(* IEC 61131-3 sources: Jacob-Formschaumtechnik-ISEL-CNC-Retrofit/twincat/PLC/src/1_IO, 3 files *)

(* ---- ST_AxisDrive.st ---- *)
(* Generische Achsschnittstelle. Die Maschinenlogik kennt nur diese Struktur.
   Die Zuordnung zu Klemmen/PDOs erfolgt ausschliesslich in FB_AxisMap_*. *)
TYPE ST_AxisDrive :
STRUCT
    (* Kommando (Logik -> Antrieb) *)
    bEnableReq   : BOOL;   (* Reglerfreigabe angefordert; wirkt nur mit Sicherheitsfreigabe *)
    bResetReq    : BOOL;
    (* Status (Antrieb -> Logik) *)
    bReady       : BOOL;
    bEnabled     : BOOL;
    bFault       : BOOL;
    nFaultCode   : UDINT;
    bHomed       : BOOL;
    bHwLimitPlus : BOOL;   (* Endschalter, Ruhestrom: FALSE = ausgeloest *)
    bHwLimitMinus: BOOL;
    rActPos      : LREAL;  (* mm *)
    rFollowErr   : LREAL;  (* mm *)
END_STRUCT
END_TYPE

(* ---- FB_AxisMap_Canopen.st ---- *)
(* Variante A: CANopen DS402 ueber EL6751. NOCH NICHT IMPLEMENTIERT.
   Wartet auf: Bestaetigung iMD 40 im Interpolated Position Mode mit TwinCAT CNC,
   PDO-Zuordnung und Achsnummern (Schaltplan fehlt). Die Logik darf diesen Baustein
   nicht direkt kennen, nur ST_AxisDrive. *)
FUNCTION_BLOCK FB_AxisMap_Canopen
VAR_INPUT
    bSafeEnable : BOOL;
END_VAR
VAR_IN_OUT
    stAxis : ST_AxisDrive;
END_VAR

(* [offen] Zuordnung der Prozessdaten *)
stAxis.bReady   := FALSE;
stAxis.bEnabled := FALSE;
stAxis.bFault   := TRUE;
stAxis.nFaultCode := 16#FFFF0001;  (* nicht implementiert: Maschine bleibt gesperrt *)
END_FUNCTION_BLOCK

(* ---- FB_AxisMap_Simulation.st ---- *)
(* Simulationsabbild fuer Usermode Runtime ohne Hardware. Folgt der Freigabe verzoegert,
   keine Bewegung. Echte Positionen kommen aus der simulierten CNC-Achse. *)
FUNCTION_BLOCK FB_AxisMap_Simulation
VAR_INPUT
    bSafeEnable : BOOL;
    bHomeReset  : BOOL;     (* Impuls: Referenzstatus loeschen *)
    bHomeCmd    : BOOL;     (* Pegel: Referenzfahrt laeuft *)
    bInjLimitPlus  : BOOL;  (* nur Simulation/Test: Endschalter Plus ausloesen *)
    bInjLimitMinus : BOOL;  (* nur Simulation/Test: Endschalter Minus ausloesen *)
    bInjFault      : BOOL;  (* nur Simulation/Test: Antriebsfehler ausloesen *)
END_VAR
VAR_IN_OUT
    stAxis : ST_AxisDrive;
END_VAR
VAR
    tonEnable : TON;
    tonHome   : TON;
END_VAR

tonEnable(IN := stAxis.bEnableReq AND bSafeEnable, PT := T#200MS);
stAxis.bReady        := TRUE;
stAxis.bEnabled      := tonEnable.Q;
stAxis.bFault        := bInjFault;
stAxis.nFaultCode    := SEL(bInjFault, 0, 16#FFFF0099);
stAxis.bHwLimitPlus  := NOT bInjLimitPlus;    (* Ruhestrom: FALSE = ausgeloest *)
stAxis.bHwLimitMinus := NOT bInjLimitMinus;

(* Referenzstatus (einzige Quelle, Befund 3): nach 2 s Referenzfahrt gesetzt, bei Reset oder Antriebsfehler geloescht *)
tonHome(IN := bHomeCmd AND stAxis.bEnabled, PT := T#2S);
IF bHomeReset OR stAxis.bFault THEN stAxis.bHomed := FALSE; END_IF
IF tonHome.Q THEN stAxis.bHomed := TRUE; END_IF
END_FUNCTION_BLOCK
